(* IEC 61131-3 sources: plc-st-coding-agent/progress/evidence/v13_rescore_20261108/candidates/codex_deepseek-v4pro, 35 files *)

(* ---- public-easy-01.st ---- *)
FUNCTION_BLOCK FB
VAR_INPUT
    bottleSensor : BOOL;
    cleaningConfirmButton : BOOL;
    fillingConfirmButton : BOOL;
    cappingConfirmButton : BOOL;
    packingConfirmButton : BOOL;
    finishedButton : BOOL;
END_VAR
VAR_OUTPUT
    Pump_Motor : BOOL;
    Filling_Valve : BOOL;
    Capping_Machine : BOOL;
    Packing_Machine : BOOL;
    Completion_Light : BOOL;
END_VAR
VAR
    cleaningConfirmEdge : BOOL;
    fillingConfirmEdge : BOOL;
    cappingConfirmEdge : BOOL;
    packingConfirmEdge : BOOL;
    finishedEdge : BOOL;
    prevCleaningConfirm : BOOL;
    prevFillingConfirm : BOOL;
    prevCappingConfirm : BOOL;
    prevPackingConfirm : BOOL;
    prevFinished : BOOL;
    CurrentStep : INT := 0;
    wasCleaning : BOOL;
END_VAR

cleaningConfirmEdge := cleaningConfirmButton AND NOT prevCleaningConfirm;
fillingConfirmEdge := fillingConfirmButton AND NOT prevFillingConfirm;
cappingConfirmEdge := cappingConfirmButton AND NOT prevCappingConfirm;
packingConfirmEdge := packingConfirmButton AND NOT prevPackingConfirm;
finishedEdge := finishedButton AND NOT prevFinished;

Pump_Motor := FALSE;
Filling_Valve := FALSE;
Capping_Machine := FALSE;
Packing_Machine := FALSE;
Completion_Light := FALSE;

IF finishedButton THEN
    IF finishedEdge THEN
        CurrentStep := 0;
    END_IF;
ELSE
    wasCleaning := (CurrentStep = 1);

    IF CurrentStep = 0 THEN
        IF bottleSensor THEN
            CurrentStep := 1;
        END_IF;
    ELSIF CurrentStep = 1 THEN
        IF cleaningConfirmEdge THEN
            CurrentStep := 2;
        END_IF;
    ELSIF CurrentStep = 2 THEN
        IF fillingConfirmEdge THEN
            CurrentStep := 3;
        END_IF;
    ELSIF CurrentStep = 3 THEN
        IF cappingConfirmEdge THEN
            CurrentStep := 4;
        END_IF;
    ELSIF CurrentStep = 4 THEN
        IF packingConfirmEdge THEN
            CurrentStep := 5;
        END_IF;
    END_IF;

    IF CurrentStep = 1 THEN
        Pump_Motor := TRUE;
    ELSIF CurrentStep = 2 THEN
        Filling_Valve := TRUE;
        IF cleaningConfirmEdge AND wasCleaning THEN
            Pump_Motor := TRUE;
        END_IF;
    ELSIF CurrentStep = 3 THEN
        Filling_Valve := TRUE;
        Capping_Machine := TRUE;
    ELSIF CurrentStep = 4 THEN
        Packing_Machine := TRUE;
    ELSIF CurrentStep = 5 THEN
        Packing_Machine := TRUE;
        Completion_Light := TRUE;
    END_IF;

    IF bottleSensor THEN
        Pump_Motor := TRUE;
    END_IF;
END_IF;

prevCleaningConfirm := cleaningConfirmButton;
prevFillingConfirm := fillingConfirmButton;
prevCappingConfirm := cappingConfirmButton;
prevPackingConfirm := packingConfirmButton;
prevFinished := finishedButton;

END_FUNCTION_BLOCK

(* ---- public-easy-02.st ---- *)
FUNCTION_BLOCK FB
VAR_INPUT
    value : DWORD;
END_VAR
VAR_OUTPUT
    hasChanged : BOOL;
    hasRisingEdges : BOOL;
    risingBits : DWORD;
    noOfRisingBits : USINT;
    hasFallingEdges : BOOL;
    fallingBits : DWORD;
    noOfFallingBits : USINT;
END_VAR
VAR
    previousValue : DWORD := 0;
    bitIndex : USINT;
END_VAR

risingBits := value AND (NOT previousValue);
fallingBits := (NOT value) AND previousValue;

noOfRisingBits := 0;
noOfFallingBits := 0;

FOR bitIndex := 0 TO 31 DO
    IF (risingBits AND SHL(DWORD#1, bitIndex)) <> 0 THEN
        noOfRisingBits := noOfRisingBits + 1;
    END_IF;
    IF (fallingBits AND SHL(DWORD#1, bitIndex)) <> 0 THEN
        noOfFallingBits := noOfFallingBits + 1;
    END_IF;
END_FOR;

hasRisingEdges := (risingBits <> 0);
hasFallingEdges := (fallingBits <> 0);
hasChanged := hasRisingEdges OR hasFallingEdges;

previousValue := value;

END_FUNCTION_BLOCK

(* ---- public-easy-03.st ---- *)
FUNCTION_BLOCK FB
VAR_INPUT
    Value      : REAL;
    hiLevel    : REAL;
    loLevel    : REAL;
    hystWindow : REAL;
END_VAR
VAR_OUTPUT
    hiAlarm : BOOL;
    loAlarm : BOOL;
    error   : BOOL;
    status  : WORD;
END_VAR
VAR
    highAlarmState : BOOL := FALSE;
    lowAlarmState  : BOOL := FALSE;
END_VAR

IF loLevel >= hiLevel THEN
    error          := TRUE;
    status         := 16#8001;
    hiAlarm        := FALSE;
    loAlarm        := FALSE;
    highAlarmState := FALSE;
    lowAlarmState  := FALSE;
ELSIF hystWindow >= (hiLevel - loLevel) THEN
    error          := TRUE;
    status         := 16#8002;
    hiAlarm        := FALSE;
    loAlarm        := FALSE;
    highAlarmState := FALSE;
    lowAlarmState  := FALSE;
ELSE
    error  := FALSE;
    status := 0;

    IF Value > hiLevel THEN
        highAlarmState := TRUE;
    ELSIF Value < (hiLevel - hystWindow) THEN
        highAlarmState := FALSE;
    END_IF;

    IF Value < loLevel THEN
        lowAlarmState := TRUE;
    ELSIF Value > (loLevel + hystWindow) THEN
        lowAlarmState := FALSE;
    END_IF;

    hiAlarm := highAlarmState;
    loAlarm := lowAlarmState;
END_IF

END_FUNCTION_BLOCK

(* ---- public-easy-04.st ---- *)
FUNCTION_BLOCK FB
VAR_INPUT
    VISCOSITY_OK : BOOL;
    PASTE_E_STOP_NC : BOOL;
    DebounceTime : TIME;
    CycleTime : TIME;
END_VAR
VAR_OUTPUT
    VFD_RUN : BOOL;
    PUMP_MAINT_DUE : BOOL;
    PUMP_RUNTIME_ACC : LINT;
END_VAR
VAR
    ViscosityValid : BOOL := FALSE;
    DebounceElapsed : TIME := T#0ms;
    RuntimeTicks : LINT := 0;
END_VAR

VFD_RUN := FALSE;

IF NOT VISCOSITY_OK THEN
    ViscosityValid := FALSE;
    DebounceElapsed := T#0ms;
ELSIF NOT PASTE_E_STOP_NC THEN
    DebounceElapsed := T#0ms;
ELSIF NOT ViscosityValid THEN
    DebounceElapsed := DebounceElapsed + CycleTime;
    IF DebounceElapsed >= DebounceTime THEN
        ViscosityValid := TRUE;
        DebounceElapsed := DebounceTime;
    END_IF
END_IF

IF PASTE_E_STOP_NC AND ViscosityValid THEN
    VFD_RUN := TRUE;
END_IF

IF VFD_RUN THEN
    RuntimeTicks := RuntimeTicks + TIME_TO_LINT(CycleTime);
END_IF

PUMP_RUNTIME_ACC := RuntimeTicks / TIME_TO_LINT(T#1h);

IF RuntimeTicks >= TIME_TO_LINT(T#500h) THEN
    PUMP_MAINT_DUE := TRUE;
ELSE
    PUMP_MAINT_DUE := FALSE;
END_IF

END_FUNCTION_BLOCK

(* ---- public-easy-05.st ---- *)
FUNCTION_BLOCK FB
VAR_INPUT
    Gap_Exceeded : BOOL;
    Weld_E_Stop_NC : BOOL;
    DebounceTime : TIME;
END_VAR
VAR_OUTPUT
    Operator_Alert : BOOL;
    Weld_Soft_Start_Active : BOOL;
END_VAR
VAR
    InitCounter : INT := 5;
    DebounceCounter : INT := 0;
END_VAR

IF InitCounter > 0 THEN
    InitCounter := InitCounter - 1;
    Weld_Soft_Start_Active := TRUE;
    Operator_Alert := FALSE;
    DebounceCounter := 0;
ELSE
    Weld_Soft_Start_Active := FALSE;

    IF NOT Weld_E_Stop_NC THEN
        Operator_Alert := FALSE;
        DebounceCounter := 0;
    ELSIF Gap_Exceeded THEN
        IF DebounceCounter < 3 THEN
            DebounceCounter := DebounceCounter + 1;
        END_IF;
        Operator_Alert := (DebounceCounter >= 3);
    ELSE
        DebounceCounter := 0;
        Operator_Alert := FALSE;
    END_IF;
END_IF;

END_FUNCTION_BLOCK

(* ---- public-easy-06.st ---- *)
FUNCTION_BLOCK FB
VAR_INPUT
    DO_LOW : BOOL;
    AERATION_E_STOP_NC : BOOL;
END_VAR
VAR_OUTPUT
    BLOWER_RUN : BOOL;
    AERATION_BLOWER_CYCLE_COUNT : UINT;
END_VAR
VAR
    first_scan : BOOL := TRUE;
    delay_counter : UINT;
    blower_run_prev : BOOL;
END_VAR

IF first_scan THEN
    BLOWER_RUN := FALSE;
    AERATION_BLOWER_CYCLE_COUNT := 0;
    delay_counter := 0;
    blower_run_prev := FALSE;
    first_scan := FALSE;
END_IF;

IF DO_LOW AND AERATION_E_STOP_NC THEN
    IF delay_counter < 5 THEN
        delay_counter := delay_counter + 1;
    END_IF;
ELSE
    delay_counter := 0;
    BLOWER_RUN := FALSE;
END_IF;

IF DO_LOW AND AERATION_E_STOP_NC AND delay_counter >= 5 THEN
    BLOWER_RUN := TRUE;
ELSE
    BLOWER_RUN := FALSE;
END_IF;

IF BLOWER_RUN AND NOT blower_run_prev THEN
    AERATION_BLOWER_CYCLE_COUNT := AERATION_BLOWER_CYCLE_COUNT + 1;
END_IF;

blower_run_prev := BLOWER_RUN;

END_FUNCTION_BLOCK

(* ---- public-hard-01.st ---- *)
FUNCTION_BLOCK FB
VAR_INPUT
    estop : BOOL;
    opeMode : BOOL;
    valveAStart : BOOL;
    valveBStart : BOOL;
    valveCStart : BOOL;
    valveDStart : BOOL;
    mixMotorStart : BOOL;
    autoStart : BOOL;
    processMode : BOOL;
    levelSensor : INT;
    mixMotorComplete : BOOL;
END_VAR
VAR_OUTPUT
    valveARun : BOOL;
    valveBRun : BOOL;
    valveCRun : BOOL;
    valveDRun : BOOL;
    mixMotorRun : BOOL;
END_VAR
VAR
    valveAStartPrev : BOOL;
    valveBStartPrev : BOOL;
    valveCStartPrev : BOOL;
    valveDStartPrev : BOOL;
    mixMotorStartPrev : BOOL;
    autoStartPrev : BOOL;
    mixMotorCompletePrev : BOOL;
    opeModePrev : BOOL;

    valveAStartR : BOOL;
    valveBStartR : BOOL;
    valveCStartR : BOOL;
    valveDStartR : BOOL;
    mixMotorStartR : BOOL;
    autoStartR : BOOL;
    mixMotorCompleteR : BOOL;
    modeChanged : BOOL;

    manualValveA : BOOL;
    manualValveB : BOOL;
    manualValveC : BOOL;
    manualValveD : BOOL;
    manualMixMotor : BOOL;

    state : INT;
    nextState : INT;
END_VAR

valveAStartR := valveAStart AND NOT valveAStartPrev;
valveBStartR := valveBStart AND NOT valveBStartPrev;
valveCStartR := valveCStart AND NOT valveCStartPrev;
valveDStartR := valveDStart AND NOT valveDStartPrev;
mixMotorStartR := mixMotorStart AND NOT mixMotorStartPrev;
autoStartR := autoStart AND NOT autoStartPrev;
mixMotorCompleteR := mixMotorComplete AND NOT mixMotorCompletePrev;
modeChanged := opeMode <> opeModePrev;

IF NOT estop THEN
    valveARun := FALSE;
    valveBRun := FALSE;
    valveCRun := FALSE;
    valveDRun := FALSE;
    mixMotorRun := FALSE;

    manualValveA := FALSE;
    manualValveB := FALSE;
    manualValveC := FALSE;
    manualValveD := FALSE;
    manualMixMotor := FALSE;
    state := 0;
    nextState := 0;

ELSIF modeChanged THEN
    valveARun := FALSE;
    valveBRun := FALSE;
    valveCRun := FALSE;
    valveDRun := FALSE;
    mixMotorRun := FALSE;

    manualValveA := FALSE;
    manualValveB := FALSE;
    manualValveC := FALSE;
    manualValveD := FALSE;
    manualMixMotor := FALSE;
    state := 0;
    nextState := 0;

ELSIF opeMode THEN
    nextState := state;

    CASE state OF
        0:
            IF autoStartR THEN
                nextState := 1;
            END_IF;

        1:
            IF levelSensor >= 50 THEN
                nextState := 2;
            END_IF;

        2:
            IF levelSensor >= 80 THEN
                IF processMode THEN
                    nextState := 3;
                ELSE
                    nextState := 4;
                END_IF;
            END_IF;

        3:
            IF levelSensor >= 100 THEN
                nextState := 4;
            END_IF;

        4:
            IF mixMotorCompleteR THEN
                nextState := 5;
            END_IF;

        5:
            IF autoStartR THEN
                nextState := 1;
            END_IF;

        ELSE
            nextState := 0;
    END_CASE;

    state := nextState;

    valveARun := FALSE;
    valveBRun := FALSE;
    valveCRun := FALSE;
    valveDRun := FALSE;
    mixMotorRun := FALSE;

    CASE state OF
        1:
            valveARun := TRUE;

        2:
            valveBRun := TRUE;

        3:
            valveCRun := TRUE;

        4:
            mixMotorRun := TRUE;

        5:
            valveDRun := TRUE;
    END_CASE;

ELSE
    IF valveAStartR THEN
        manualValveA := NOT manualValveA;
    END_IF;

    IF valveBStartR THEN
        manualValveB := NOT manualValveB;
    END_IF;

    IF valveCStartR THEN
        manualValveC := NOT manualValveC;
    END_IF;

    IF valveDStartR THEN
        manualValveD := NOT manualValveD;
    END_IF;

    IF mixMotorStartR THEN
        manualMixMotor := NOT manualMixMotor;
    END_IF;

    valveARun := manualValveA;
    valveBRun := manualValveB;
    valveCRun := manualValveC;
    valveDRun := manualValveD;
    mixMotorRun := manualMixMotor;
END_IF;

valveAStartPrev := valveAStart;
valveBStartPrev := valveBStart;
valveCStartPrev := valveCStart;
valveDStartPrev := valveDStart;
mixMotorStartPrev := mixMotorStart;
autoStartPrev := autoStart;
mixMotorCompletePrev := mixMotorComplete;
opeModePrev := opeMode;

END_FUNCTION_BLOCK

(* ---- public-hard-02.st ---- *)
FUNCTION_BLOCK FB
VAR_INPUT
    processLength : USINT;
    sensor1 : BOOL;
    sensor2 : BOOL;
    sensor3 : BOOL;
    sensor4 : BOOL;
    sensor5 : BOOL;
    station1Start : BOOL;
    station2Complete : BOOL;
    station3Complete : BOOL;
    station4Complete : BOOL;
    processSequence : ARRAY[1..8] OF USINT;
END_VAR
VAR_OUTPUT
    conveyorLeft : BOOL;
    conveyorRight : BOOL;
END_VAR
VAR
    phase : USINT := 0;
    curStation : USINT := 1;
    dstStation : USINT := 0;
    idx : USINT := 0;
    startEdge : BOOL;
    station2Edge : BOOL;
    station3Edge : BOOL;
    station4Edge : BOOL;
    compEdge : BOOL;
    lastStation1Start : BOOL;
    lastStation2Complete : BOOL;
    lastStation3Complete : BOOL;
    lastStation4Complete : BOOL;
END_VAR

startEdge := station1Start AND NOT lastStation1Start;
station2Edge := station2Complete AND NOT lastStation2Complete;
station3Edge := station3Complete AND NOT lastStation3Complete;
station4Edge := station4Complete AND NOT lastStation4Complete;

compEdge := FALSE;
IF phase = 2 THEN
    IF curStation = 2 THEN
        compEdge := station2Edge;
    ELSIF curStation = 3 THEN
        compEdge := station3Edge;
    ELSIF curStation = 4 THEN
        compEdge := station4Edge;
    END_IF;
END_IF;

IF phase = 0 THEN
    IF startEdge AND sensor1 THEN
        IF processLength >= 1 AND processLength <= 8 THEN
            idx := 1;
            dstStation := processSequence[1];
            phase := 1;
        END_IF;
    END_IF;
ELSIF phase = 1 THEN
    IF dstStation = 2 AND sensor2 THEN
        curStation := 2;
        phase := 2;
    ELSIF dstStation = 3 AND sensor3 THEN
        curStation := 3;
        phase := 2;
    ELSIF dstStation = 4 AND sensor4 THEN
        curStation := 4;
        phase := 2;
    ELSIF dstStation = 5 AND sensor5 THEN
        curStation := 5;
        phase := 0;
    END_IF;
ELSIF phase = 2 THEN
    IF compEdge THEN
        idx := idx + 1;
        IF idx <= processLength THEN
            dstStation := processSequence[idx];
            IF dstStation = curStation THEN
                phase := 2;
            ELSE
                phase := 1;
            END_IF;
        ELSE
            phase := 0;
        END_IF;
    END_IF;
END_IF;

conveyorLeft := FALSE;
conveyorRight := FALSE;
IF phase = 1 THEN
    IF dstStation > curStation THEN
        conveyorRight := TRUE;
    ELSIF dstStation < curStation THEN
        conveyorLeft := TRUE;
    END_IF;
END_IF;

lastStation1Start := station1Start;
lastStation2Complete := station2Complete;
lastStation3Complete := station3Complete;
lastStation4Complete := station4Complete;

END_FUNCTION_BLOCK

(* ---- public-hard-03.st ---- *)
FUNCTION_BLOCK FB
VAR_INPUT
    addRecipe : BOOL;
    deleteRecipe : BOOL;
    modifyRecipe : BOOL;
    queryRecipe : BOOL;
    recipeIn : ST_Recipe;
END_VAR
VAR_OUTPUT
    recipeAdded : BOOL;
    recipeDeleted : BOOL;
    recipeModified : BOOL;
    recipeQueryResult : ST_Recipe;
    error : BOOL;
    status : WORD;
END_VAR
VAR_IN_OUT
    recipe : ARRAY[1..10] OF ST_Recipe;
END_VAR
VAR
    lastAddRecipe : BOOL;
    lastDeleteRecipe : BOOL;
    lastModifyRecipe : BOOL;
    lastQueryRecipe : BOOL;
    addEdge : BOOL;
    deleteEdge : BOOL;
    modifyEdge : BOOL;
    queryEdge : BOOL;
    i : INT;
    foundIndex : INT;
    emptyIndex : INT;
    recipeFound : BOOL;
END_VAR

recipeAdded := FALSE;
recipeDeleted := FALSE;
recipeModified := FALSE;

addEdge := addRecipe AND NOT lastAddRecipe;
deleteEdge := deleteRecipe AND NOT lastDeleteRecipe;
modifyEdge := modifyRecipe AND NOT lastModifyRecipe;
queryEdge := queryRecipe AND NOT lastQueryRecipe;

IF addEdge OR deleteEdge OR modifyEdge OR queryEdge THEN
    error := FALSE;
    status := WORD#0;
END_IF

IF queryEdge THEN
    recipeFound := FALSE;
    foundIndex := 0;

    FOR i := 1 TO 10 DO
        IF (recipeIn.recipeID <> 0) AND (recipe[i].recipeID = recipeIn.recipeID) THEN
            recipeFound := TRUE;
            foundIndex := i;
        END_IF
    END_FOR

    IF recipeFound THEN
        recipeQueryResult := recipe[foundIndex];
    ELSE
        error := TRUE;
        status := WORD#16#8001;
        recipeQueryResult.recipeID := 0;
        recipeQueryResult.ingredientType := 0;
        recipeQueryResult.ingredientRatio := 0.0;
        recipeQueryResult.productionTemperature := 0.0;
    END_IF
END_IF

IF addEdge THEN
    recipeFound := FALSE;
    emptyIndex := 0;

    FOR i := 1 TO 10 DO
        IF recipe[i].recipeID = recipeIn.recipeID THEN
            recipeFound := TRUE;
        END_IF

        IF (recipe[i].recipeID = 0) AND (emptyIndex = 0) THEN
            emptyIndex := i;
        END_IF
    END_FOR

    IF recipeFound THEN
        error := TRUE;
        status := WORD#16#8002;
    ELSIF emptyIndex = 0 THEN
        error := TRUE;
        status := WORD#16#8003;
    ELSE
        recipe[emptyIndex] := recipeIn;
        recipeAdded := TRUE;
    END_IF
END_IF

IF deleteEdge THEN
    recipeFound := FALSE;
    foundIndex := 0;

    FOR i := 1 TO 10 DO
        IF (recipeIn.recipeID <> 0) AND (recipe[i].recipeID = recipeIn.recipeID) THEN
            recipeFound := TRUE;
            foundIndex := i;
        END_IF
    END_FOR

    IF recipeFound THEN
        recipe[foundIndex].recipeID := 0;
        recipeDeleted := TRUE;
    ELSE
        error := TRUE;
        status := WORD#16#8004;
    END_IF
END_IF

IF modifyEdge THEN
    recipeFound := FALSE;
    foundIndex := 0;

    FOR i := 1 TO 10 DO
        IF (recipeIn.recipeID <> 0) AND (recipe[i].recipeID = recipeIn.recipeID) THEN
            recipeFound := TRUE;
            foundIndex := i;
        END_IF
    END_FOR

    IF recipeFound THEN
        recipe[foundIndex] := recipeIn;
        recipeModified := TRUE;
    ELSE
        error := TRUE;
        status := WORD#16#8005;
    END_IF
END_IF

lastAddRecipe := addRecipe;
lastDeleteRecipe := deleteRecipe;
lastModifyRecipe := modifyRecipe;
lastQueryRecipe := queryRecipe;
END_FUNCTION_BLOCK

(* ---- public-hard-04.st ---- *)
FUNCTION_BLOCK FB
VAR_INPUT
    enqueue : BOOL;
    dequeue : BOOL;
    reset : BOOL;
    capacity : DINT;
END_VAR
VAR_OUTPUT
    elementCount : DINT;
    status : WORD;
END_VAR
VAR_IN_OUT
    item : DINT;
    buffer : ARRAY[1..4] OF DINT;
END_VAR
VAR
    head : DINT := 1;
    tail : DINT := 1;
    count : DINT := 0;
    prevEnqueue : BOOL := FALSE;
    prevDequeue : BOOL := FALSE;
    enqRise : BOOL := FALSE;
    deqRise : BOOL := FALSE;
END_VAR

elementCount := count;
status := 16#0000;

enqRise := enqueue AND NOT prevEnqueue;
deqRise := dequeue AND NOT prevDequeue;

IF reset THEN
    count := 0;
    head := 1;
    tail := 1;
    elementCount := count;
ELSIF NOT (enqRise AND deqRise) THEN
    IF enqRise THEN
        IF count < capacity THEN
            buffer[tail] := item;
            tail := tail + 1;
            IF tail > capacity THEN
                tail := 1;
            END_IF
            count := count + 1;
        ELSE
            status := 16#8002;
        END_IF
    END_IF

    IF deqRise THEN
        IF count > 0 THEN
            item := buffer[head];
            head := head + 1;
            IF head > capacity THEN
                head := 1;
            END_IF
            count := count - 1;
        ELSE
            status := 16#8001;
        END_IF
    END_IF

    elementCount := count;
END_IF

prevEnqueue := enqueue;
prevDequeue := dequeue;

END_FUNCTION_BLOCK

(* ---- public-hard-05.st ---- *)
FUNCTION_BLOCK FB
VAR_INPUT
    ManualMode : BOOL;
    SingleStepMode : BOOL;
    SingleCycleMode : BOOL;
    ContinuousMode : BOOL;
    EmergencyStop : BOOL;
    Start : BOOL;
    DownButton : BOOL;
    UpButton : BOOL;
    LeftButton : BOOL;
    RightButton : BOOL;
    GripButton : BOOL;
    ReleaseButton : BOOL;
    DownLimitSwitch : BOOL;
    UpLimitSwitch : BOOL;
    LeftLimitSwitch : BOOL;
    RightLimitSwitch : BOOL;
    GripLimitSwitch : BOOL;
    ReleaseLimitSwitch : BOOL;
END_VAR
VAR_OUTPUT
    MoveDown : BOOL;
    MoveUp : BOOL;
    MoveLeft : BOOL;
    MoveRight : BOOL;
    ActivateGrip : BOOL;
    ActivateRelease : BOOL;
END_VAR
VAR
    StartPrev : BOOL;
    StartPulse : BOOL;
    ModeId : INT;
    PrevModeId : INT;
    Step : INT := 0;
    StepDone : BOOL;
    WDown : BOOL;
    WUp : BOOL;
    WLeft : BOOL;
    WRight : BOOL;
    WGrip : BOOL;
    WRelease : BOOL;
    AutoDown : BOOL;
    AutoUp : BOOL;
    AutoLeft : BOOL;
    AutoRight : BOOL;
    AutoGrip : BOOL;
    AutoRelease : BOOL;
END_VAR

StartPulse := Start AND NOT StartPrev;
StartPrev := Start;

IF ManualMode THEN
    ModeId := 1;
ELSIF SingleStepMode THEN
    ModeId := 2;
ELSIF SingleCycleMode THEN
    ModeId := 3;
ELSIF ContinuousMode THEN
    ModeId := 4;
ELSE
    ModeId := 0;
END_IF

IF ModeId <> PrevModeId THEN
    Step := 0;
END_IF
PrevModeId := ModeId;

StepDone := FALSE;
CASE Step OF
    1: StepDone := DownLimitSwitch;
    2: StepDone := GripLimitSwitch;
    3: StepDone := UpLimitSwitch;
    4: StepDone := RightLimitSwitch;
    5: StepDone := DownLimitSwitch;
    6: StepDone := ReleaseLimitSwitch;
    7: StepDone := UpLimitSwitch;
    8: StepDone := LeftLimitSwitch;
END_CASE

IF EmergencyStop THEN
    IF ModeId = 2 THEN
        IF StartPulse THEN
            IF Step = 0 THEN
                Step := 1;
            ELSIF StepDone THEN
                IF Step = 8 THEN
                    Step := 1;
                ELSE
                    Step := Step + 1;
                END_IF
            END_IF
        END_IF
    ELSIF ModeId = 3 THEN
        IF StartPulse AND (Step = 0) THEN
            Step := 1;
        ELSIF (Step > 0) AND StepDone THEN
            IF Step = 8 THEN
                Step := 0;
            ELSE
                Step := Step + 1;
            END_IF
        END_IF
    ELSIF ModeId = 4 THEN
        IF StartPulse AND (Step = 0) THEN
            Step := 1;
        ELSIF (Step > 0) AND StepDone THEN
            IF Step = 8 THEN
                Step := 1;
            ELSE
                Step := Step + 1;
            END_IF
        END_IF
    END_IF
END_IF

AutoDown := FALSE;
AutoUp := FALSE;
AutoLeft := FALSE;
AutoRight := FALSE;
AutoGrip := FALSE;
AutoRelease := FALSE;

CASE Step OF
    1: AutoDown := NOT DownLimitSwitch;
    2: AutoGrip := NOT GripLimitSwitch;
    3: AutoUp := NOT UpLimitSwitch;
    4: AutoRight := NOT RightLimitSwitch;
    5: AutoDown := NOT DownLimitSwitch;
    6: AutoRelease := NOT ReleaseLimitSwitch;
    7: AutoUp := NOT UpLimitSwitch;
    8: AutoLeft := NOT LeftLimitSwitch;
END_CASE

IF EmergencyStop THEN
    IF ModeId = 1 THEN
        WDown := DownButton AND NOT DownLimitSwitch;
        WUp := UpButton AND NOT UpLimitSwitch AND NOT WDown;
        WLeft := LeftButton AND NOT LeftLimitSwitch;
        WRight := RightButton AND NOT RightLimitSwitch AND NOT WLeft;
        WGrip := GripButton AND NOT GripLimitSwitch;
        WRelease := ReleaseButton AND NOT ReleaseLimitSwitch AND NOT WGrip;
    ELSIF (ModeId = 2) OR (ModeId = 3) OR (ModeId = 4) THEN
        WDown := AutoDown;
        WUp := AutoUp;
        WLeft := AutoLeft;
        WRight := AutoRight;
        WGrip := AutoGrip;
        WRelease := AutoRelease;
    ELSE
        WDown := FALSE;
        WUp := FALSE;
        WLeft := FALSE;
        WRight := FALSE;
        WGrip := FALSE;
        WRelease := FALSE;
    END_IF
ELSE
    WDown := FALSE;
    WUp := FALSE;
    WLeft := FALSE;
    WRight := FALSE;
    WGrip := FALSE;
    WRelease := FALSE;
END_IF

MoveDown := WDown;
MoveUp := WUp;
MoveLeft := WLeft;
MoveRight := WRight;
ActivateGrip := WGrip;
ActivateRelease := WRelease;
END_FUNCTION_BLOCK

(* ---- public-hard-06.st ---- *)
FUNCTION_BLOCK FB
VAR_INPUT
    Mode : BOOL;
    ForwardButton : BOOL;
    ReverseButton : BOOL;
    SensorFeed : BOOL;
    SensorWash : BOOL;
    SensorWeight : BOOL;
    SensorFiring : BOOL;
    SensorOutput : BOOL;
    washComplete : BOOL;
    weightComplete : BOOL;
    weight : REAL;
    firingComplete : BOOL;
END_VAR
VAR_OUTPUT
    MotorForward : BOOL;
    MotorReverse : BOOL;
    kick : BOOL;
    CompletionLight : BOOL;
    firingTemp : REAL;
END_VAR
VAR
    AutoState : INT := 0;
    washPrev : BOOL;
    weightPrev : BOOL;
    firingPrev : BOOL;
    washRising : BOOL;
    weightRising : BOOL;
    firingRising : BOOL;
    tempCalc : REAL := 0.0;
END_VAR

washRising := washComplete AND NOT washPrev;
weightRising := weightComplete AND NOT weightPrev;
firingRising := firingComplete AND NOT firingPrev;

kick := FALSE;

IF Mode THEN
    CASE AutoState OF
        0:
            IF SensorOutput THEN
                AutoState := 8;
            ELSIF SensorFiring THEN
                AutoState := 6;
            ELSIF SensorWeight THEN
                AutoState := 4;
            ELSIF SensorWash THEN
                AutoState := 2;
            ELSIF SensorFeed THEN
                AutoState := 1;
            END_IF;

        1:
            IF SensorWash THEN
                AutoState := 2;
            END_IF;

        2:
            IF washRising THEN
                AutoState := 3;
            END_IF;

        3:
            IF SensorWeight THEN
                AutoState := 4;
            END_IF;

        4:
            IF NOT SensorWeight THEN
                AutoState := 0;
            ELSIF weightRising THEN
                IF (weight >= 100.0) AND (weight <= 200.0) THEN
                    tempCalc := 500.0 + (weight - 100.0) * 0.5;
                    AutoState := 5;
                ELSE
                    tempCalc := 0.0;
                END_IF;
            END_IF;

        5:
            IF SensorFiring THEN
                AutoState := 6;
            END_IF;

        6:
            IF firingRising THEN
                AutoState := 7;
            END_IF;

        7:
            IF SensorOutput THEN
                AutoState := 8;
            END_IF;

        8:
            IF NOT SensorOutput THEN
                AutoState := 0;
            END_IF;
    END_CASE;

    IF (AutoState = 4) AND weightRising AND ((weight < 100.0) OR (weight > 200.0)) THEN
        kick := TRUE;
    END_IF;

    MotorForward := (AutoState = 1) OR (AutoState = 3) OR (AutoState = 5) OR (AutoState = 7);
    MotorReverse := FALSE;
ELSE
    AutoState := 0;
    MotorForward := ForwardButton AND NOT ReverseButton;
    MotorReverse := ReverseButton AND NOT ForwardButton;
END_IF

washPrev := washComplete;
weightPrev := weightComplete;
firingPrev := firingComplete;

CompletionLight := SensorOutput;
firingTemp := tempCalc;

(* ---- public-medium-01.st ---- *)
TYPE ST_Pump :
STRUCT
    priority : INT;
    selection : BOOL;
    RunComd : BOOL;
END_STRUCT
END_TYPE

FUNCTION_BLOCK FB
VAR_INPUT
    mode : BOOL;
    start : BOOL;
    stop : BOOL;
END_VAR
VAR_IN_OUT
    pumpGroup : ARRAY[1..5] OF ST_Pump;
END_VAR
VAR
    i : INT;
    pass : INT;
    bestIdx : INT;
    maxP : INT;
    selected : ARRAY[1..5] OF BOOL;
END_VAR

FOR i := 1 TO 5 DO
    selected[i] := FALSE;
END_FOR

IF mode AND start AND NOT stop THEN
    FOR pass := 1 TO 3 DO
        bestIdx := 0;
        maxP := -32768;
        FOR i := 1 TO 5 DO
            IF NOT selected[i] THEN
                IF bestIdx = 0 THEN
                    bestIdx := i;
                    maxP := pumpGroup[i].priority;
                ELSIF pumpGroup[i].priority > maxP THEN
                    bestIdx := i;
                    maxP := pumpGroup[i].priority;
                END_IF
            END_IF
        END_FOR
        IF bestIdx <> 0 THEN
            selected[bestIdx] := TRUE;
        END_IF
    END_FOR
END_IF

FOR i := 1 TO 5 DO
    IF stop THEN
        pumpGroup[i].RunComd := FALSE;
    ELSIF NOT start THEN
        pumpGroup[i].RunComd := FALSE;
    ELSIF mode THEN
        pumpGroup[i].RunComd := selected[i];
    ELSE
        pumpGroup[i].RunComd := pumpGroup[i].selection;
    END_IF
END_FOR

END_FUNCTION_BLOCK

(* ---- public-medium-02.st ---- *)
TYPE ST_AnalogChannel :
STRUCT
    enable : BOOL;
    hiLIM : REAL;
    loLIM : REAL;
    bipolar : BOOL;
    measuringMode : INT;
    retVal : WORD;
    outputValue : REAL;
END_STRUCT
END_TYPE

FUNCTION_BLOCK FB
VAR_INPUT
    count : DINT;
END_VAR
VAR_IN_OUT
    analogValues : ARRAY[1..8] OF INT;
    channels : ARRAY[1..8] OF ST_AnalogChannel;
END_VAR
VAR
    idx : DINT;
    rawValue : REAL;
    scalingSpan : REAL;
END_VAR

IF count >= 1 THEN
    FOR idx := 1 TO count DO
        IF channels[idx].enable THEN
            channels[idx].retVal := 0;

            IF (channels[idx].measuringMode < 0) OR (channels[idx].measuringMode > 2) THEN
                channels[idx].retVal := 16#8001;
            ELSIF channels[idx].hiLIM <= channels[idx].loLIM THEN
                channels[idx].retVal := 16#8002;
            ELSE
                rawValue := INT_TO_REAL(analogValues[idx]);

                IF channels[idx].measuringMode = 0 THEN
                    scalingSpan := channels[idx].hiLIM - channels[idx].loLIM;

                    IF channels[idx].bipolar THEN
                        channels[idx].outputValue := channels[idx].loLIM
                            + ((rawValue + 27648.0) * scalingSpan / 55296.0);
                    ELSE
                        channels[idx].outputValue := channels[idx].loLIM
                            + (rawValue * scalingSpan / 27648.0);
                    END_IF;

                ELSIF channels[idx].measuringMode = 1 THEN
                    channels[idx].outputValue := rawValue / 10.0;

                ELSE
                    channels[idx].outputValue := rawValue / 100.0;
                END_IF;
            END_IF;
        END_IF;
    END_FOR;
END_IF;

END_FUNCTION_BLOCK

(* ---- public-medium-03.st ---- *)
FUNCTION_BLOCK FB
VAR_INPUT
    cyclicExecution : BOOL;
    trigger : BOOL;
    value : LREAL;
    windowSize : INT;
    reset : BOOL;
END_VAR
VAR_OUTPUT
    average : LREAL;
    windowSizeReached : BOOL;
    error : BOOL;
    status : WORD;
END_VAR
VAR
    samples : ARRAY[0..99] OF LREAL;
    sampleCount : INT := 0;
    sum : LREAL := 0.0;
    triggerOld : BOOL;
    triggerRising : BOOL;
    i : INT;
    j : INT;
END_VAR

triggerRising := trigger AND NOT triggerOld;

IF windowSize < 1 OR windowSize > 100 THEN
    IF reset THEN
        sampleCount := 0;
        sum := 0.0;
    END_IF

    error := TRUE;
    status := 16#8200;
    average := 0.0;
    windowSizeReached := FALSE;
ELSE
    error := FALSE;
    status := 16#0000;

    IF reset THEN
        sampleCount := 0;
        sum := 0.0;
        average := 0.0;
        windowSizeReached := FALSE;
    ELSE
        IF sampleCount > windowSize THEN
            j := 0;
            FOR i := sampleCount - windowSize TO sampleCount - 1 DO
                samples[j] := samples[i];
                j := j + 1;
            END_FOR
            sampleCount := windowSize;
        END_IF

        IF cyclicExecution OR triggerRising THEN
            IF sampleCount < windowSize THEN
                samples[sampleCount] := value;
                sampleCount := sampleCount + 1;
            ELSE
                IF windowSize > 1 THEN
                    FOR i := 0 TO windowSize - 2 DO
                        samples[i] := samples[i + 1];
                    END_FOR
                END_IF
                samples[windowSize - 1] := value;
            END_IF
        END_IF

        sum := 0.0;
        IF sampleCount > 0 THEN
            FOR i := 0 TO sampleCount - 1 DO
                sum := sum + samples[i];
            END_FOR
            average := sum / INT_TO_LREAL(sampleCount);
            windowSizeReached := sampleCount >= windowSize;
        ELSE
            average := 0.0;
            windowSizeReached := FALSE;
        END_IF
    END_IF
END_IF

triggerOld := trigger;

END_FUNCTION_BLOCK

(* ---- public-medium-04.st ---- *)
FUNCTION_BLOCK FB
VAR_INPUT
    TemperatureSensorInput: REAL;
    SetTemperature: REAL;
END_VAR
VAR_OUTPUT
    CurrentTemperature: REAL;
    SetTempDisplay: REAL;
    HeaterStatus: BOOL;
    OverheatProtection: BOOL;
    HeaterOutput: BOOL;
END_VAR
VAR
    HeatRunCounter: INT := 0;
    OverheatRemaining: INT := 0;
    SensorFault: BOOL;
END_VAR

CurrentTemperature := TemperatureSensorInput;
SetTempDisplay := SetTemperature;
SensorFault := TemperatureSensorInput < 0.0 OR TemperatureSensorInput > 100.0;

IF OverheatRemaining > 0 THEN
    OverheatProtection := TRUE;
    HeaterOutput := FALSE;
    HeatRunCounter := 0;
    OverheatRemaining := OverheatRemaining - 1;
ELSIF SensorFault THEN
    OverheatProtection := FALSE;
    HeaterOutput := FALSE;
    HeatRunCounter := 0;
ELSIF TemperatureSensorInput >= SetTemperature THEN
    OverheatProtection := FALSE;
    HeaterOutput := FALSE;
    HeatRunCounter := 0;
ELSIF TemperatureSensorInput < SetTemperature THEN
    OverheatProtection := FALSE;
    HeaterOutput := TRUE;
    HeatRunCounter := HeatRunCounter + 1;

    IF HeatRunCounter >= 5 THEN
        HeaterOutput := FALSE;
        OverheatProtection := TRUE;
        HeatRunCounter := 0;
        OverheatRemaining := 2;
    END_IF
END_IF

HeaterStatus := HeaterOutput;

END_FUNCTION_BLOCK

(* ---- public-medium-05.st ---- *)
FUNCTION_BLOCK FB
VAR_INPUT
    Mode : BOOL;
    ForwardButton : BOOL;
    ReverseButton : BOOL;
    SensorA : BOOL;
    SensorB : BOOL;
    SensorC : BOOL;
    ButtonA : BOOL;
    ButtonB : BOOL;
    ButtonC : BOOL;
END_VAR
VAR_OUTPUT
    MotorForward : BOOL;
    MotorReverse : BOOL;
    CompletionLight : BOOL;
END_VAR
VAR
    ButtonA_Prev : BOOL;
    ButtonB_Prev : BOOL;
    ButtonC_Prev : BOOL;
    ButtonA_Rising : BOOL;
    ButtonB_Rising : BOOL;
    ButtonC_Rising : BOOL;
    MovingAB : BOOL;
    MovingBC : BOOL;
    WorkComplete : BOOL;
END_VAR

MotorForward := FALSE;
MotorReverse := FALSE;
CompletionLight := FALSE;

ButtonA_Rising := ButtonA AND NOT ButtonA_Prev;
ButtonB_Rising := ButtonB AND NOT ButtonB_Prev;
ButtonC_Rising := ButtonC AND NOT ButtonC_Prev;

IF NOT Mode THEN
    MovingAB := FALSE;
    MovingBC := FALSE;
    WorkComplete := FALSE;

    IF ForwardButton AND NOT ReverseButton THEN
        MotorForward := TRUE;
    END_IF;

    IF ReverseButton AND NOT ForwardButton THEN
        MotorReverse := TRUE;
    END_IF;
ELSE
    IF SensorB AND MovingAB THEN
        MovingAB := FALSE;
    END_IF;

    IF SensorC AND MovingBC THEN
        MovingBC := FALSE;
    END_IF;

    IF NOT SensorC THEN
        WorkComplete := FALSE;
    END_IF;

    IF SensorA AND ButtonA_Rising AND NOT MovingAB AND NOT MovingBC THEN
        MovingAB := TRUE;
    END_IF;

    IF SensorB AND ButtonB_Rising AND NOT MovingBC THEN
        MovingBC := TRUE;
    END_IF;

    IF SensorC AND ButtonC_Rising THEN
        WorkComplete := TRUE;
    END_IF;

    MotorForward := MovingAB OR MovingBC;
    CompletionLight := SensorC AND WorkComplete;
END_IF;

ButtonA_Prev := ButtonA;
ButtonB_Prev := ButtonB;
ButtonC_Prev := ButtonC;
END_FUNCTION_BLOCK

(* ---- public-medium-06.st ---- *)
FUNCTION_BLOCK FB
VAR_INPUT
    THICKNESS_FAULT : BOOL;
    THICKNESS_SIGNAL_VALID : BOOL;
    CUTTING_RUN : BOOL;
    FaultTimestamp : DINT;
    CycleTime : TIME;
END_VAR
VAR_OUTPUT
    THICKNESS_ALARM : BOOL;
    Slab_Fault_Counter : UINT;
    Slab_Runtime_Accumulator : LINT;
    Slab_Fault_History : ARRAY[0..4] OF DINT;
END_VAR
VAR
    PreviousValidFault : BOOL := FALSE;
    AlarmHoldActive : BOOL := FALSE;
    AlarmHoldElapsed : TIME := T#0MS;
    HistoryIndex : INT;
END_VAR

IF NOT THICKNESS_SIGNAL_VALID THEN
    THICKNESS_ALARM := FALSE;
    AlarmHoldActive := FALSE;
    AlarmHoldElapsed := T#0MS;
    PreviousValidFault := FALSE;
ELSE
    IF THICKNESS_FAULT AND NOT PreviousValidFault THEN
        Slab_Fault_Counter := Slab_Fault_Counter + UINT#1;

        FOR HistoryIndex := 4 TO 1 BY -1 DO
            Slab_Fault_History[HistoryIndex] := Slab_Fault_History[HistoryIndex - 1];
        END_FOR;

        Slab_Fault_History[0] := FaultTimestamp;
        AlarmHoldActive := TRUE;
        AlarmHoldElapsed := T#0MS;
    END_IF;

    IF THICKNESS_FAULT THEN
        THICKNESS_ALARM := TRUE;
        AlarmHoldActive := TRUE;
    ELSE
        IF AlarmHoldActive AND (AlarmHoldElapsed < T#500MS) THEN
            THICKNESS_ALARM := TRUE;
        ELSE
            THICKNESS_ALARM := FALSE;
            AlarmHoldActive := FALSE;
            AlarmHoldElapsed := T#0MS;
        END_IF;
    END_IF;

    IF AlarmHoldActive AND (AlarmHoldElapsed < T#500MS) THEN
        AlarmHoldElapsed := AlarmHoldElapsed + CycleTime;
    END_IF;

    PreviousValidFault := THICKNESS_FAULT;

    IF CUTTING_RUN AND NOT THICKNESS_FAULT THEN
        Slab_Runtime_Accumulator := Slab_Runtime_Accumulator + TIME_TO_LINT(CycleTime);
    END_IF;
END_IF;
END_FUNCTION_BLOCK

(* ---- public-medium-07.st ---- *)
FUNCTION_BLOCK FB
VAR_INPUT
    OCCUPANCY_DETECTED : BOOL;
    ENERGY_SAVING_MODE : BOOL;
    HVAC_MODE_SELECTOR : INT;
END_VAR
VAR_OUTPUT
    SUPPLY_FAN_RUN : BOOL;
    TEMP_SETPOINT_ADJUST : INT;
END_VAR
VAR
    FanStartCounter : DINT := 0;
END_VAR

SUPPLY_FAN_RUN := FALSE;
TEMP_SETPOINT_ADJUST := 0;

IF OCCUPANCY_DETECTED AND HVAC_MODE_SELECTOR <> 3 THEN
    FanStartCounter := FanStartCounter + 1;
    IF FanStartCounter >= 30 THEN
        SUPPLY_FAN_RUN := TRUE;
    END_IF;
ELSE
    FanStartCounter := 0;
    SUPPLY_FAN_RUN := FALSE;
END_IF;

CASE HVAC_MODE_SELECTOR OF
    0:
        IF OCCUPANCY_DETECTED THEN
            TEMP_SETPOINT_ADJUST := 0;
        ELSIF ENERGY_SAVING_MODE THEN
            TEMP_SETPOINT_ADJUST := 3;
        ELSE
            TEMP_SETPOINT_ADJUST := 2;
        END_IF;

    1:
        IF OCCUPANCY_DETECTED THEN
            TEMP_SETPOINT_ADJUST := 0;
        ELSE
            TEMP_SETPOINT_ADJUST := 1;
        END_IF;

    2:
        IF OCCUPANCY_DETECTED THEN
            TEMP_SETPOINT_ADJUST := 0;
        ELSE
            TEMP_SETPOINT_ADJUST := 4;
        END_IF;

    3:
        TEMP_SETPOINT_ADJUST := 4;

    ELSE
        TEMP_SETPOINT_ADJUST := 0;
END_CASE;

IF TEMP_SETPOINT_ADJUST > 4 THEN
    TEMP_SETPOINT_ADJUST := 4;
ELSIF TEMP_SETPOINT_ADJUST < -4 THEN
    TEMP_SETPOINT_ADJUST := -4;
END_IF;

END_FUNCTION_BLOCK

(* ---- public-medium-08.st ---- *)
FUNCTION_BLOCK FB
VAR_INPUT
    ipText : STRING(254);
END_VAR
VAR_OUTPUT
    ipValue : UDINT;
END_VAR
VAR
    scanIndex : INT;
    currentChar : STRING(1);
    currentSegment : UDINT;
    digitValue : UDINT;
    segmentCount : INT;
    hasDigit : BOOL;
    isValid : BOOL;
    ok : BOOL;
END_VAR

ipValue := UDINT#0;
currentSegment := UDINT#0;
segmentCount := 0;
hasDigit := FALSE;
isValid := TRUE;

FOR scanIndex := 1 TO LEN(ipText) BY 1 DO
    IF isValid THEN
        currentChar := MID(ipText, 1, scanIndex);

        IF currentChar = '.' THEN
            IF hasDigit THEN
                segmentCount := segmentCount + 1;
                ipValue := (ipValue * UDINT#256) + currentSegment;
                currentSegment := UDINT#0;
                hasDigit := FALSE;
            ELSE
                isValid := FALSE;
            END_IF
        ELSIF currentChar = '0' THEN
            digitValue := UDINT#0;
            hasDigit := TRUE;
            currentSegment := (currentSegment * UDINT#10) + digitValue;
            IF currentSegment > UDINT#255 THEN
                isValid := FALSE;
            END_IF
        ELSIF currentChar = '1' THEN
            digitValue := UDINT#1;
            hasDigit := TRUE;
            currentSegment := (currentSegment * UDINT#10) + digitValue;
            IF currentSegment > UDINT#255 THEN
                isValid := FALSE;
            END_IF
        ELSIF currentChar = '2' THEN
            digitValue := UDINT#2;
            hasDigit := TRUE;
            currentSegment := (currentSegment * UDINT#10) + digitValue;
            IF currentSegment > UDINT#255 THEN
                isValid := FALSE;
            END_IF
        ELSIF currentChar = '3' THEN
            digitValue := UDINT#3;
            hasDigit := TRUE;
            currentSegment := (currentSegment * UDINT#10) + digitValue;
            IF currentSegment > UDINT#255 THEN
                isValid := FALSE;
            END_IF
        ELSIF currentChar = '4' THEN
            digitValue := UDINT#4;
            hasDigit := TRUE;
            currentSegment := (currentSegment * UDINT#10) + digitValue;
            IF currentSegment > UDINT#255 THEN
                isValid := FALSE;
            END_IF
        ELSIF currentChar = '5' THEN
            digitValue := UDINT#5;
            hasDigit := TRUE;
            currentSegment := (currentSegment * UDINT#10) + digitValue;
            IF currentSegment > UDINT#255 THEN
                isValid := FALSE;
            END_IF
        ELSIF currentChar = '6' THEN
            digitValue := UDINT#6;
            hasDigit := TRUE;
            currentSegment := (currentSegment * UDINT#10) + digitValue;
            IF currentSegment > UDINT#255 THEN
                isValid := FALSE;
            END_IF
        ELSIF currentChar = '7' THEN
            digitValue := UDINT#7;
            hasDigit := TRUE;
            currentSegment := (currentSegment * UDINT#10) + digitValue;
            IF currentSegment > UDINT#255 THEN
                isValid := FALSE;
            END_IF
        ELSIF currentChar = '8' THEN
            digitValue := UDINT#8;
            hasDigit := TRUE;
            currentSegment := (currentSegment * UDINT#10) + digitValue;
            IF currentSegment > UDINT#255 THEN
                isValid := FALSE;
            END_IF
        ELSIF currentChar = '9' THEN
            digitValue := UDINT#9;
            hasDigit := TRUE;
            currentSegment := (currentSegment * UDINT#10) + digitValue;
            IF currentSegment > UDINT#255 THEN
                isValid := FALSE;
            END_IF
        ELSE
            isValid := FALSE;
        END_IF
    END_IF
END_FOR

IF isValid THEN
    IF hasDigit THEN
        segmentCount := segmentCount + 1;
        ipValue := (ipValue * UDINT#256) + currentSegment;
    ELSE
        isValid := FALSE;
    END_IF
END_IF

IF isValid AND (segmentCount <> 4) THEN
    isValid := FALSE;
END_IF

IF isValid THEN
    ok := TRUE;
ELSE
    ipValue := UDINT#0;
    ok := FALSE;
END_IF

END_FUNCTION_BLOCK

(* ---- self-easy-01.st ---- *)
FUNCTION_BLOCK FB
VAR_INPUT
    enable : BOOL;
    values : ARRAY[1..8] OF INT;
    count : INT;
    avgEnable : BOOL;
END_VAR
VAR_OUTPUT
    avgOut : REAL;
END_VAR
VAR
    lastAvg : REAL := 0.0;
    total : LINT;
    sampleCount : INT;
    i : INT;
    avg : REAL;
END_VAR

avgOut := lastAvg;

IF enable AND avgEnable AND (count > 0) THEN
    sampleCount := count;
    IF sampleCount > 8 THEN
        sampleCount := 8;
    END_IF;

    total := 0;
    FOR i := 1 TO sampleCount DO
        total := total + INT_TO_LINT(values[i]);
    END_FOR;

    avg := LINT_TO_REAL(total) / INT_TO_REAL(sampleCount);
    avgOut := avg;
    lastAvg := avg;
END_IF;

END_FUNCTION_BLOCK

(* ---- self-easy-02.st ---- *)
FUNCTION_BLOCK FB
VAR_INPUT
    tankLevel : REAL;
    outletFlow : REAL;
    inletPermit : BOOL;
    resetBtn : BOOL;
END_VAR
VAR_OUTPUT
    pumpRun : BOOL;
    alarmHigh : BOOL;
    alarmLow : BOOL;
    outletValveOpen : BOOL;
END_VAR
VAR
    resetBtnPrev : BOOL := FALSE;
    resetRising : BOOL;
    highLatched : BOOL := FALSE;
    lowLatched : BOOL := FALSE;
END_VAR

resetRising := resetBtn AND NOT resetBtnPrev;

IF tankLevel >= 85.0 THEN
    highLatched := TRUE;
END_IF

IF tankLevel <= 15.0 THEN
    lowLatched := TRUE;
END_IF

IF resetRising THEN
    IF tankLevel < 85.0 THEN
        highLatched := FALSE;
    END_IF
    IF tankLevel > 15.0 THEN
        lowLatched := FALSE;
    END_IF
END_IF

alarmHigh := highLatched;
alarmLow := lowLatched;

IF inletPermit AND NOT highLatched AND tankLevel >= 15.0 AND tankLevel < 85.0 THEN
    pumpRun := TRUE;
ELSE
    pumpRun := FALSE;
END_IF

IF NOT lowLatched AND tankLevel > 15.0 THEN
    outletValveOpen := TRUE;
ELSE
    outletValveOpen := FALSE;
END_IF

resetBtnPrev := resetBtn;

END_FUNCTION_BLOCK

(* ---- self-hard-01.st ---- *)
FUNCTION_BLOCK FB
VAR_INPUT
    flowLow : BOOL;
    ackBtn : BOOL;
    sensorOK : BOOL;
END_VAR
VAR_OUTPUT
    alarmActive : BOOL;
    alarmAcked : BOOL;
    highHigh : BOOL;
END_VAR
VAR
    lastAck : BOOL := FALSE;
    lastFlow : BOOL := FALSE;
    ackRise : BOOL;
    flowRise : BOOL;
    activeState : BOOL := FALSE;
    ackState : BOOL := FALSE;
END_VAR

ackRise := ackBtn AND NOT lastAck;
flowRise := flowLow AND NOT lastFlow;

IF ackRise THEN
    IF flowLow THEN
        activeState := TRUE;
        ackState := TRUE;
    ELSE
        activeState := FALSE;
        ackState := FALSE;
    END_IF;
ELSIF flowRise THEN
    activeState := TRUE;
    ackState := FALSE;
ELSIF flowLow THEN
    activeState := TRUE;
ELSE
    IF NOT activeState THEN
        activeState := FALSE;
        ackState := FALSE;
    ELSIF NOT ackState THEN
        activeState := TRUE;
        ackState := TRUE;
    ELSE
        activeState := FALSE;
        ackState := FALSE;
    END_IF;
END_IF;

alarmActive := activeState;
alarmAcked := ackState;
highHigh := NOT sensorOK;

lastAck := ackBtn;
lastFlow := flowLow;
END_FUNCTION_BLOCK

(* ---- self-hard-02.st ---- *)
FUNCTION_BLOCK FB
VAR_INPUT
    startBtn : BOOL;
    abortBtn : BOOL;
    setpoint : REAL;
    pv : REAL;
    maxDuration : INT;
END_VAR
VAR_OUTPUT
    elapsed : INT;
    phase : INT;
    timeout : BOOL;
END_VAR
VAR
    startRising : BOOL;
    lastStart : BOOL;
END_VAR

startRising := startBtn AND NOT lastStart;

IF startRising THEN
    elapsed := 0;
    phase := 1;
    timeout := FALSE;
ELSIF abortBtn THEN
    phase := 9;
ELSIF (phase = 1) OR (phase = 2) THEN
    elapsed := elapsed + 1;

    IF elapsed >= maxDuration THEN
        timeout := TRUE;
        phase := 3;
    ELSIF (phase = 1) AND (pv >= setpoint) THEN
        phase := 2;
    END_IF;
END_IF;

lastStart := startBtn;
END_FUNCTION_BLOCK

(* ---- self-hard-03.st ---- *)
FUNCTION_BLOCK FB
VAR_INPUT
    pushEn   : BOOL;
    pushItem : INT;
    popEn    : BOOL;
END_VAR
VAR_OUTPUT
    count  : INT;
    full   : BOOL;
    empty  : BOOL;
    head   : INT;
END_VAR
VAR_IN_OUT
    fifo : ARRAY[1..8] OF INT;
END_VAR
VAR
    pushPrev : BOOL;
    popPrev  : BOOL;
    pushRise : BOOL;
    popRise  : BOOL;
    i        : INT;
END_VAR

pushRise := pushEn AND NOT pushPrev;
popRise  := popEn AND NOT popPrev;
pushPrev := pushEn;
popPrev  := popEn;

IF popRise THEN
    IF count > 0 THEN
        FOR i := 1 TO 7 DO
            fifo[i] := fifo[i + 1];
        END_FOR;
        fifo[8] := 0;
        count := count - 1;
    END_IF;
END_IF;

IF pushRise THEN
    IF count < 8 THEN
        fifo[count + 1] := pushItem;
        count := count + 1;
    END_IF;
END_IF;

full := count >= 8;
empty := count <= 0;

IF count <= 0 THEN
    head := 0;
ELSE
    head := fifo[1];
END_IF;

END_FUNCTION_BLOCK

(* ---- self-hard-04.st ---- *)
FUNCTION_BLOCK FB
VAR_INPUT
    demand : INT;
    runHours : ARRAY[1..5] OF LINT;
    rotated : BOOL;
END_VAR
VAR_OUTPUT
    leadPump : INT;
    lagPump : INT;
    runningCount : INT;
END_VAR
VAR
    clipped : INT;
    order : ARRAY[1..5] OF INT;
    i : INT;
    j : INT;
    tempIdx : INT;
    bestLead : INT;
    bestLag : INT;
    currentLeadHours : LINT;
    bestLeadHours : LINT;
    memLead : INT := 0;
    memLag : INT := 0;
END_VAR

clipped := demand;
IF clipped < 0 THEN
    clipped := 0;
ELSIF clipped > 5 THEN
    clipped := 5;
END_IF

runningCount := clipped;

IF clipped = 0 THEN
    memLead := 0;
    memLag := 0;
ELSE
    order[1] := 1;
    order[2] := 2;
    order[3] := 3;
    order[4] := 4;
    order[5] := 5;

    FOR i := 1 TO 4 DO
        FOR j := i + 1 TO 5 DO
            IF (runHours[order[j]] < runHours[order[i]]) OR ((runHours[order[j]] = runHours[order[i]]) AND (order[j] < order[i])) THEN
                tempIdx := order[i];
                order[i] := order[j];
                order[j] := tempIdx;
            END_IF
        END_FOR
    END_FOR

    bestLead := order[1];
    IF clipped >= 2 THEN
        bestLag := order[2];
    ELSE
        bestLag := 0;
    END_IF

    IF memLead = 0 THEN
        memLead := bestLead;
        memLag := bestLag;
    ELSE
        IF rotated THEN
            currentLeadHours := runHours[memLead];
            bestLeadHours := runHours[bestLead];
            IF (bestLead <> memLead) AND ((currentLeadHours - bestLeadHours) > 50) THEN
                memLead := bestLead;
                IF clipped >= 2 THEN
                    memLag := bestLag;
                ELSE
                    memLag := 0;
                END_IF
            END_IF
        END_IF

        IF clipped >= 2 THEN
            IF (memLag = 0) OR (memLag = memLead) THEN
                memLag := 0;
                FOR i := 1 TO 5 DO
                    IF (order[i] <> memLead) AND (memLag = 0) THEN
                        memLag := order[i];
                    END_IF
                END_FOR
            END_IF
        ELSE
            memLag := 0;
        END_IF
    END_IF
END_IF

leadPump := memLead;
lagPump := memLag;
END_FUNCTION_BLOCK

(* ---- self-hard-05.st ---- *)
FUNCTION_BLOCK FB
VAR_INPUT
    runRequest : BOOL;
    flameOK : BOOL;
    o2Valid : BOOL;
    o2PV : REAL;
    baseAir : REAL;
    resetBtn : BOOL;
END_VAR
VAR_OUTPUT
    fuelPermit : BOOL;
    trimEnable : BOOL;
    airTrim : REAL;
    airCommand : REAL;
    tripLatched : BOOL;
    o2Fault : BOOL;
END_VAR
VAR
    prevResetBtn : BOOL := FALSE;
END_VAR

o2Fault := (NOT o2Valid) OR (o2PV < 0.0) OR (o2PV > 21.0);

IF runRequest AND (NOT flameOK) THEN
    tripLatched := TRUE;
ELSIF tripLatched AND resetBtn AND (NOT prevResetBtn)
      AND (NOT runRequest) AND (NOT flameOK) THEN
    tripLatched := FALSE;
END_IF;

prevResetBtn := resetBtn;

fuelPermit := runRequest AND flameOK AND (NOT tripLatched);

trimEnable := fuelPermit AND (NOT o2Fault);

IF trimEnable THEN
    airTrim := 2.0 * (2.0 - o2PV);
    IF airTrim < -10.0 THEN
        airTrim := -10.0;
    END_IF;
    IF airTrim > 10.0 THEN
        airTrim := 10.0;
    END_IF;
ELSE
    airTrim := 0.0;
END_IF;

IF fuelPermit THEN
    airCommand := baseAir + airTrim;
    IF airCommand < 0.0 THEN
        airCommand := 0.0;
    END_IF;
    IF airCommand > 100.0 THEN
        airCommand := 100.0;
    END_IF;
ELSE
    airCommand := 0.0;
END_IF;

END_FUNCTION_BLOCK

(* ---- self-hard-06.st ---- *)
FUNCTION_BLOCK FB
VAR_INPUT
    runRequest : BOOL;
    pressure : REAL;
    pressureValid : BOOL;
    fuelFlow : REAL;
    steamFlow : REAL;
    outletCmd : INT;
    outletFeedback : INT;
    resetBtn : BOOL;
END_VAR
VAR_OUTPUT
    tripLatched : BOOL;
    fuelPermit : BOOL;
    currentCauseMask : WORD;
    latchedCauseMask : WORD;
    diagnosticActive : BOOL;
END_VAR
VAR
    resetBtnPrev : BOOL;
    resetRising : BOOL;
    valveStuckCnt : INT;
END_VAR

resetRising := resetBtn AND NOT resetBtnPrev;

IF runRequest AND pressureValid AND (pressure >= 4500.0)
   AND (outletCmd >= 50) AND (outletFeedback <= 10) THEN
    valveStuckCnt := valveStuckCnt + 1;
ELSE
    valveStuckCnt := 0;
END_IF

currentCauseMask := 0;

IF runRequest THEN
    IF NOT pressureValid THEN
        currentCauseMask := currentCauseMask OR WORD#16#0001;
    ELSIF pressure >= 4500.0 THEN
        IF valveStuckCnt >= 3 THEN
            currentCauseMask := currentCauseMask OR WORD#16#0002;
        END_IF
        IF fuelFlow >= 4.0 AND steamFlow <= 10.0 THEN
            currentCauseMask := currentCauseMask OR WORD#16#0004;
        END_IF
        IF currentCauseMask = 0 THEN
            currentCauseMask := WORD#16#0008;
        END_IF
    END_IF
END_IF

IF runRequest AND (NOT pressureValid OR pressure >= 4500.0) THEN
    tripLatched := TRUE;
ELSIF resetRising AND NOT runRequest AND pressureValid AND pressure <= 4200.0 THEN
    tripLatched := FALSE;
    latchedCauseMask := 0;
END_IF

IF tripLatched THEN
    latchedCauseMask := latchedCauseMask OR currentCauseMask;
END_IF

fuelPermit := runRequest AND NOT tripLatched;
diagnosticActive := currentCauseMask <> 0;

resetBtnPrev := resetBtn;

END_FUNCTION_BLOCK

(* ---- self-hard-07.st ---- *)
FUNCTION_BLOCK FB
VAR_INPUT
    mode : INT;
    resetBtn : BOOL;
    scanSeconds : REAL;
    tempSP : REAL;
    tempPV : REAL;
    flowPV : REAL;
    manualFlowSP : REAL;
    manualValve : REAL;
END_VAR
VAR_OUTPUT
    flowSP : REAL;
    valveCommand : REAL;
    fault : BOOL;
    normalMode : BOOL;
END_VAR
VAR
    initialized : BOOL;
    prevMode : INT;
    prevReset : BOOL;
    prevFlowSP : REAL;
    prevValveCommand : REAL;

    resetRising : BOOL;
    modeChanged : BOOL;
    outerIntegral : REAL;
    innerIntegral : REAL;
    tempError : REAL;
    flowError : REAL;
    rawOutput : REAL;
END_VAR

fault := (mode < 0) OR (mode > 2)
         OR (scanSeconds <= 0.0)
         OR (scanSeconds > 10.0);

resetRising := resetBtn AND (NOT prevReset);

IF NOT initialized THEN
    normalMode := FALSE;
    flowSP := manualFlowSP;
    valveCommand := manualValve;
    outerIntegral := flowSP - 1.0 * (tempSP - tempPV);
    innerIntegral := valveCommand - 2.0 * (flowSP - flowPV);
ELSIF fault THEN
    normalMode := FALSE;
    flowSP := manualFlowSP;
    valveCommand := manualValve;
    outerIntegral := flowSP - 1.0 * (tempSP - tempPV);
    innerIntegral := valveCommand - 2.0 * (flowSP - flowPV);
ELSIF resetRising THEN
    normalMode := FALSE;
    flowSP := manualFlowSP;
    valveCommand := manualValve;
    outerIntegral := flowSP - 1.0 * (tempSP - tempPV);
    innerIntegral := valveCommand - 2.0 * (flowSP - flowPV);
ELSE
    modeChanged := mode <> prevMode;

    IF modeChanged THEN
        normalMode := FALSE;
        valveCommand := prevValveCommand;

        IF mode = 2 THEN
            flowSP := prevFlowSP;
        ELSE
            flowSP := manualFlowSP;
        END_IF;

        outerIntegral := flowSP - 1.0 * (tempSP - tempPV);
        innerIntegral := valveCommand - 2.0 * (flowSP - flowPV);
    ELSE
        normalMode := TRUE;

        IF mode = 0 THEN
            flowSP := manualFlowSP;
            valveCommand := manualValve;
            outerIntegral := flowSP - 1.0 * (tempSP - tempPV);
            innerIntegral := valveCommand - 2.0 * (flowSP - flowPV);
        ELSIF mode = 1 THEN
            flowSP := manualFlowSP;
            outerIntegral := flowSP - 1.0 * (tempSP - tempPV);

            flowError := flowSP - flowPV;
            innerIntegral := innerIntegral + 0.5 * flowError * scanSeconds;
            rawOutput := 2.0 * flowError + innerIntegral;

            IF rawOutput < 0.0 THEN
                valveCommand := 0.0;
            ELSIF rawOutput > 100.0 THEN
                valveCommand := 100.0;
            ELSE
                valveCommand := rawOutput;
            END_IF;

            innerIntegral := valveCommand - 2.0 * flowError;
        ELSE
            tempError := tempSP - tempPV;
            outerIntegral := outerIntegral + 0.2 * tempError * scanSeconds;
            rawOutput := 1.0 * tempError + outerIntegral;

            IF rawOutput < 0.0 THEN
                flowSP := 0.0;
            ELSIF rawOutput > 50.0 THEN
                flowSP := 50.0;
            ELSE
                flowSP := rawOutput;
            END_IF;

            outerIntegral := flowSP - 1.0 * tempError;

            flowError := flowSP - flowPV;
            innerIntegral := innerIntegral + 0.5 * flowError * scanSeconds;
            rawOutput := 2.0 * flowError + innerIntegral;

            IF rawOutput < 0.0 THEN
                valveCommand := 0.0;
            ELSIF rawOutput > 100.0 THEN
                valveCommand := 100.0;
            ELSE
                valveCommand := rawOutput;
            END_IF;

            innerIntegral := valveCommand - 2.0 * flowError;
        END_IF;
    END_IF;
END_IF;

prevFlowSP := flowSP;
prevValveCommand := valveCommand;
prevMode := mode;
prevReset := resetBtn;
initialized := TRUE;

END_FUNCTION_BLOCK

(* ---- self-medium-01.st ---- *)
TYPE ST_Recipe :
STRUCT
    recipeID : INT;
    totalRatio : REAL;
    temperature : REAL;
END_STRUCT
END_TYPE

FUNCTION_BLOCK FB
VAR_INPUT
    recipe : ARRAY[1..8] OF ST_Recipe;
    selSlot : INT;
    loadCmd : BOOL;
    running : BOOL;
END_VAR
VAR_OUTPUT
    valid : BOOL;
    loadedID : INT;
END_VAR
VAR
    lastLoadCmd : BOOL;
    loadRising : BOOL;
    slotValid : BOOL;
END_VAR

loadRising := loadCmd AND NOT lastLoadCmd;
slotValid := (selSlot >= 1) AND (selSlot <= 8);

IF running THEN
    valid := FALSE;
ELSIF loadRising THEN
    IF NOT slotValid THEN
        valid := FALSE;
        loadedID := 0;
    ELSIF recipe[selSlot].recipeID = 0 THEN
        valid := FALSE;
    ELSIF (recipe[selSlot].totalRatio < 99.0) OR (recipe[selSlot].totalRatio > 101.0) THEN
        valid := FALSE;
        loadedID := 0;
    ELSIF (recipe[selSlot].temperature < 30.0) OR (recipe[selSlot].temperature > 180.0) THEN
        valid := FALSE;
        loadedID := 0;
    ELSE
        valid := TRUE;
        loadedID := recipe[selSlot].recipeID;
    END_IF
END_IF

lastLoadCmd := loadCmd;

END_FUNCTION_BLOCK

(* ---- self-medium-02.st ---- *)
FUNCTION_BLOCK FB
VAR_INPUT
    enable : BOOL;
    rawValue : REAL;
END_VAR
VAR_OUTPUT
    filteredValue : REAL;
    windowFull : BOOL;
    sampleCount : INT;
END_VAR
VAR
    buffer : ARRAY[0..7] OF REAL;
    writeIndex : INT := 0;
    validCount : INT := 0;
    sum : REAL;
    i : INT;
END_VAR

IF enable THEN
    buffer[writeIndex] := rawValue;

    writeIndex := writeIndex + 1;
    IF writeIndex >= 8 THEN
        writeIndex := 0;
    END_IF;

    IF validCount < 8 THEN
        validCount := validCount + 1;
    END_IF;

    sum := 0.0;
    FOR i := 0 TO validCount - 1 DO
        sum := sum + buffer[i];
    END_FOR;

    filteredValue := sum / INT_TO_REAL(validCount);
    sampleCount := validCount;
    windowFull := validCount >= 8;
ELSE
    validCount := 0;
    writeIndex := 0;
    sampleCount := 0;
    windowFull := FALSE;
END_IF;

END_FUNCTION_BLOCK

(* ---- self-medium-03.st ---- *)
FUNCTION_BLOCK FB
VAR_INPUT
    openBtn    : BOOL;
    closeBtn   : BOOL;
    openLimit  : BOOL;
    closeLimit : BOOL;
    obstacle   : BOOL;
END_VAR
VAR_OUTPUT
    motorUp   : BOOL;
    motorDown : BOOL;
    errorFlag : BOOL;
END_VAR
VAR
    state        : INT := 0; (* 0=IDLE, 1=OPENING, 2=CLOSING, 3=FAULT *)
    openBtnPrev  : BOOL := FALSE;
    closeBtnPrev : BOOL := FALSE;
    bothPrev     : BOOL := FALSE;
    openBtnRise  : BOOL;
    closeBtnRise : BOOL;
    bothPressed  : BOOL;
    resetRise    : BOOL;
END_VAR

openBtnRise  := openBtn AND NOT openBtnPrev;
closeBtnRise := closeBtn AND NOT closeBtnPrev;
bothPressed  := openBtn AND closeBtn;
resetRise    := bothPressed AND NOT bothPrev;

CASE state OF
    0: (* IDLE *)
        motorUp   := FALSE;
        motorDown := FALSE;
        errorFlag := FALSE;

        IF openBtnRise AND NOT openLimit THEN
            state := 1;
        ELSIF closeBtnRise AND NOT closeLimit THEN
            state := 2;
        END_IF;

    1: (* OPENING *)
        IF obstacle THEN
            motorUp   := FALSE;
            motorDown := FALSE;
            errorFlag := TRUE;
            state     := 3;
        ELSIF openLimit THEN
            motorUp   := FALSE;
            motorDown := FALSE;
            errorFlag := FALSE;
            state     := 0;
        ELSE
            motorUp   := TRUE;
            motorDown := FALSE;
            errorFlag := FALSE;
        END_IF;

    2: (* CLOSING *)
        IF obstacle THEN
            motorDown := FALSE;
            errorFlag := FALSE;
            state     := 1;

            IF openLimit THEN
                motorUp := FALSE;
            ELSE
                motorUp := TRUE;
            END_IF;
        ELSIF closeLimit THEN
            motorUp   := FALSE;
            motorDown := FALSE;
            errorFlag := FALSE;
            state     := 0;
        ELSE
            motorUp   := FALSE;
            motorDown := TRUE;
            errorFlag := FALSE;
        END_IF;

    3: (* FAULT *)
        motorUp   := FALSE;
        motorDown := FALSE;
        errorFlag := TRUE;

        IF resetRise AND NOT obstacle THEN
            errorFlag := FALSE;
            state     := 0;
        END_IF;
END_CASE;

openBtnPrev  := openBtn;
closeBtnPrev := closeBtn;
bothPrev     := bothPressed;
END_FUNCTION_BLOCK

(* ---- self-medium-04.st ---- *)
FUNCTION_BLOCK FB
VAR_INPUT
    startBtn : BOOL;
    resetBtn : BOOL;
    doneSensor : BOOL;
    targetVol : REAL;
    flowVol : REAL;
END_VAR
VAR_OUTPUT
    valveOpen : BOOL;
    fillsToday : INT;
END_VAR
VAR
    startR : BOOL;
    resetR : BOOL;
    lastStart : BOOL;
    lastReset : BOOL;
    accumulated : REAL;
    stage : INT;
END_VAR

startR := startBtn AND NOT lastStart;
resetR := resetBtn AND NOT lastReset;

IF resetR THEN
    stage := 0;
    valveOpen := FALSE;
    fillsToday := 0;
    accumulated := 0.0;
ELSIF startR AND stage = 0 THEN
    stage := 1;
    valveOpen := TRUE;
    accumulated := 0.0;
END_IF;

IF stage = 1 THEN
    accumulated := accumulated + flowVol;
    IF accumulated >= targetVol THEN
        valveOpen := FALSE;
        stage := 2;
    END_IF;
END_IF;

IF stage = 2 AND doneSensor THEN
    fillsToday := fillsToday + 1;
    stage := 0;
END_IF;

lastStart := startBtn;
lastReset := resetBtn;

END_FUNCTION_BLOCK

(* ---- self-medium-05.st ---- *)
FUNCTION_BLOCK FB
VAR_INPUT
    enable : BOOL;
    resetBtn : BOOL;
    scanSeconds : LREAL;
    steamFlow : LREAL;
    fuelFlow : LREAL;
    steamTemp : LREAL;
    steamPressure : LREAL;
END_VAR
VAR_OUTPUT
    qualified : BOOL;
    dataFault : BOOL;
    qualifiedTon : LREAL;
    fuelTon : LREAL;
    revenue : LREAL;
    cost : LREAL;
    netProfit : LREAL;
END_VAR
VAR
    prevResetBtn : BOOL;
END_VAR

qualified := (steamTemp >= 447.0) AND (steamTemp <= 453.0)
             AND (steamPressure >= 3750.0) AND (steamPressure <= 3850.0);

dataFault := (scanSeconds <= 0.0) OR (scanSeconds > 10.0)
             OR (steamFlow < 0.0) OR (steamFlow > 90.0)
             OR (fuelFlow < 0.0) OR (fuelFlow > 6.0);

IF resetBtn AND NOT prevResetBtn THEN
    qualifiedTon := 0.0;
    fuelTon := 0.0;
ELSE
    IF enable AND NOT dataFault THEN
        IF qualified THEN
            qualifiedTon := qualifiedTon + steamFlow * scanSeconds / 1000.0;
        END_IF;

        fuelTon := fuelTon + fuelFlow * scanSeconds / 1000.0;
    END_IF;
END_IF;

prevResetBtn := resetBtn;

revenue := qualifiedTon * 280.0;
cost := fuelTon * 1500.0;
netProfit := revenue - cost;

END_FUNCTION_BLOCK

(* ---- self-medium-06.st ---- *)
FUNCTION_BLOCK FB
VAR_INPUT
    enable : BOOL;
    resetBtn : BOOL;
    sensorValid : BOOL;
    setpoint : REAL;
    temperature : REAL;
    scanSeconds : REAL;
    bias : REAL;
END_VAR
VAR_OUTPUT
    power : REAL;
    correction : REAL;
    fault : BOOL;
END_VAR
VAR
    resetPrev : BOOL;
    resetRising : BOOL;
    ePrev : REAL;
    bHist : BOOL;
    e : REAL;
    de : REAL;
    x : REAL;
    y : REAL;
    muNx : REAL;
    muZx : REAL;
    muPx : REAL;
    muNy : REAL;
    muZy : REAL;
    muPy : REAL;
    w : REAL;
    num : REAL;
    den : REAL;
    rawPower : REAL;
END_VAR

resetRising := resetBtn AND NOT resetPrev;
resetPrev := resetBtn;

fault := (NOT sensorValid) OR (scanSeconds <= 0.0) OR (scanSeconds > 10.0);

IF (NOT enable) OR resetRising OR fault THEN
    power := 0.0;
    correction := 0.0;
    ePrev := 0.0;
    bHist := FALSE;
ELSE
    e := setpoint - temperature;

    IF bHist THEN
        de := (e - ePrev) / scanSeconds;
    ELSE
        de := 0.0;
    END_IF;

    x := e / 10.0;
    IF x < -1.0 THEN
        x := -1.0;
    ELSIF x > 1.0 THEN
        x := 1.0;
    END_IF;

    y := de / 2.0;
    IF y < -1.0 THEN
        y := -1.0;
    ELSIF y > 1.0 THEN
        y := 1.0;
    END_IF;

    muNx := -x;
    IF muNx < 0.0 THEN
        muNx := 0.0;
    END_IF;

    IF x >= 0.0 THEN
        muZx := 1.0 - x;
    ELSE
        muZx := 1.0 + x;
    END_IF;

    muPx := x;
    IF muPx < 0.0 THEN
        muPx := 0.0;
    END_IF;

    muNy := -y;
    IF muNy < 0.0 THEN
        muNy := 0.0;
    END_IF;

    IF y >= 0.0 THEN
        muZy := 1.0 - y;
    ELSE
        muZy := 1.0 + y;
    END_IF;

    muPy := y;
    IF muPy < 0.0 THEN
        muPy := 0.0;
    END_IF;

    num := 0.0;
    den := 0.0;

    w := muNx;
    IF muNy < w THEN
        w := muNy;
    END_IF;
    num := num + w * (-30.0);
    den := den + w;

    w := muNx;
    IF muZy < w THEN
        w := muZy;
    END_IF;
    num := num + w * (-20.0);
    den := den + w;

    w := muNx;
    IF muPy < w THEN
        w := muPy;
    END_IF;
    num := num + w * (-10.0);
    den := den + w;

    w := muZx;
    IF muNy < w THEN
        w := muNy;
    END_IF;
    num := num + w * (-10.0);
    den := den + w;

    w := muZx;
    IF muZy < w THEN
        w := muZy;
    END_IF;
    num := num + w * 0.0;
    den := den + w;

    w := muZx;
    IF muPy < w THEN
        w := muPy;
    END_IF;
    num := num + w * 10.0;
    den := den + w;

    w := muPx;
    IF muNy < w THEN
        w := muNy;
    END_IF;
    num := num + w * 10.0;
    den := den + w;

    w := muPx;
    IF muZy < w THEN
        w := muZy;
    END_IF;
    num := num + w * 20.0;
    den := den + w;

    w := muPx;
    IF muPy < w THEN
        w := muPy;
    END_IF;
    num := num + w * 30.0;
    den := den + w;

    IF den > 0.0 THEN
        correction := num / den;
    ELSE
        correction := 0.0;
    END_IF;

    rawPower := bias + correction;
    IF rawPower < 0.0 THEN
        power := 0.0;
    ELSIF rawPower > 100.0 THEN
        power := 100.0;
    ELSE
        power := rawPower;
    END_IF;

    ePrev := e;
    bHist := TRUE;
END_IF;

END_FUNCTION_BLOCK
